(* PLC project PLC_ST_Auto, PLC_ST_Auto 1.0 *)
(* stored: creationDateTime 2026-11-09T06:11:21 *)

PROGRAM DualMotorSequentialStart
  VAR_INPUT
    start : BOOL;
    stop : BOOL;
  END_VAR
  VAR_OUTPUT
    motor1 : BOOL;
    motor2 : BOOL;
  END_VAR
  VAR
    run_latch : BOOL;
    delay_tmr : TON;
  END_VAR

      (* Assumption: stop is a normally-open button (TRUE = pressed). *)
(* Start/stop latch with stop dominant *)
run_latch := (start OR run_latch) AND NOT stop;

(* Motor1 starts immediately when latched *)
motor1 := run_latch;

(* Motor2 starts after 3 s of motor1 running *)
delay_tmr(IN := run_latch, PT := T#3s);
motor2 := delay_tmr.Q AND run_latch;
    
END_PROGRAM

CONFIGURATION Config
  RESOURCE Res ON PLC
    TASK MainTask(INTERVAL := T#10ms, PRIORITY := 1);
    PROGRAM DualMotorSequentialStart_inst WITH MainTask : DualMotorSequentialStart;
  END_RESOURCE
END_CONFIGURATION
